(* IEC 61131-3 sources: Lasal-MCP/examples/SampleSource/LASALScreenAdvancedSolution/LASALScreenAdvancedSolution/LASALScreenAdvacnedSolution/Stations/Terminal/HMI/Class/CirleMyIO, 1 file *)

(* ---- CirleMyIO.st ---- *)
(*!
<Class
	Name               = "CirleMyIO"
	Revision           = "0.0"
	RealtimeTask       = "false"
	CyclicTask         = "false"
	BackgroundTask     = "false"
	Sigmatek           = "false"
	OSInterface        = "false"
	HighPriority       = "false"
	Automatic          = "false"
	UpdateMode         = "Prescan"
	SharedCommandTable = "true"
	Objectsize         = "(510,660)">
	<Channels>
		<Server Name="CircleAngle" Visualized="true" Initialize="true" DefValue="3600" WriteProtected="false" Retentive="File"/>
		<Server Name="CircleRadius" Visualized="true" Initialize="true" DefValue="80" WriteProtected="false" Retentive="File"/>
		<Server Name="XPos" Visualized="true" Initialize="true" DefValue="60" WriteProtected="false" Retentive="false"/>
		<Server Name="YPos" Visualized="true" Initialize="true" DefValue="60" WriteProtected="false" Retentive="false"/>
		<Client Name="_Grafix" Required="false" Internal="false"/>
	</Channels>
	<Network Name="CirleMyIO">
		<!-- List of Components in this network -->
		<Components>
			<Object
				Name       = "_base"
				Class      = "_MyIO"
				Position   = "(218,120)"
				Visualized = "true"
				Remotely   = "true">
				<Channels>
					<Server Name="Refresh"/>
					<Server Name="Server0"/>
					<Client Name="Graphic"/>
					<Client Name="Lse"/>
				</Channels>
			</Object>
		</Components>
		<Comments>
		</Comments>
		<!-- List of Connections in this network -->
		<Connections>
			<Connection Source="this.Server0" Destination="_base.Server0" Vertices="(706,210),(534,210),"/>
			<Connection Source="this.Refresh" Destination="_base.Refresh" Vertices="(706,270),(534,270),"/>
			<Connection Source="_base.Lse" Destination="this.Lse" Vertices="(218,210),(38,210),"/>
		</Connections>
		<!-- Headerfiles -->
		<Options>
		</Options>
	</Network>
</Class>
*)
#pragma using _MyIO

CirleMyIO : CLASS
: _MyIO
  //Servers:
	XPos 	: SvrCh_DINT;
	YPos 	: SvrCh_DINT;
	CircleRadius 	: SvrCh_DINT;
	CircleAngle 	: SvrCh_DINT;
  //Clients:
	_Grafix 	: CltChCmd__Grafix;
  //Variables:
		myFocus 	: BOOL;
		TempX 	: _KOORD;
		TempY 	: _KOORD;
  //Functions:
				//! <Function Comment="this method will be called once when the focus will be given to this object" Name="GetFocus"/>
	FUNCTION __CDECL VIRTUAL GLOBAL GetFocus
		VAR_INPUT
			pio 	: ^_IO;			//! <Variable Comment="pointer to _IO information" Name="GetFocus.pio"/>
		END_VAR
		VAR_OUTPUT
			retcode (EAX) 	: _DOIT;			//! <Variable Comment="return _IFAILED if you dont want to get the focus on the other hand _IDLE" Name="GetFocus.retcode"/>
		END_VAR;
				//! <Function Comment="this method is called once when the focus is taken from object" Name="KillFocus"/>
	FUNCTION __CDECL VIRTUAL GLOBAL KillFocus
		VAR_INPUT
			pio 	: ^_IO;			//! <Variable Comment="pointer to _IO information" Name="KillFocus.pio"/>
		END_VAR
		VAR_OUTPUT
			retcode (EAX) 	: _DOIT;			//! <Variable Comment="return always _IDLE because you can&apos;t prevent action" Name="KillFocus.retcode"/>
		END_VAR;
				//! <Function Comment="this method is called everytime when the input is active and a event occured" Name="GetEvent"/>
	FUNCTION __CDECL VIRTUAL GLOBAL GetEvent
		VAR_INPUT
			ped 	: ^_EDITOR;			//! <Variable Comment="pointer to _EDITOR information" Name="GetEvent.ped"/>
			pe 	: ^_EVENT;			//! <Variable Comment="pointer to _EVENT information" Name="GetEvent.pe"/>
		END_VAR
		VAR_OUTPUT
			retcode (EAX) 	: _DOIT;			//! <Variable Comment="for the returnstatement there are 3 different possibilities&#13;&#10;  _IDLE ..... the system should goon like it is (system goes on)&#13;&#10;  _IDIDIT ... i did it (system is ready)&#13;&#10;  _IFAILED .. i tried to do my best, but i failed (system is ready)&#13;&#10;" Name="GetEvent.retcode"/>
		END_VAR;
				//! <Function Comment="this method is called everytime when system wants to redraw the io" Name="Draw"/>
	FUNCTION __CDECL VIRTUAL GLOBAL Draw
		VAR_INPUT
			pio 	: ^_IO;			//! <Variable Comment="pointer to _IO information" Name="Draw.pio"/>
			pr 	: ^_RESULT;			//! <Variable Comment="pointer to _RESULT information" Name="Draw.pr"/>
			pv 	: ^_VARIABLE;			//! <Variable Comment="pointer to io _VARIABLE information" Name="Draw.pv"/>
			input 	: BOOL;			//! <Variable Comment="TRUE it&apos;s an input&#13;&#10;FALSE it&apos;s an output" Name="Draw.input"/>
		END_VAR
		VAR_OUTPUT
			retcode (EAX) 	: _DOIT;			//! <Variable Comment="for the returnstatement there are 3 different possibilities&#13;&#10;  _IDLE ..... the system should goon like it is (system goes on)&#13;&#10;  _IDIDIT ... i did it (system is ready)&#13;&#10;  _IFAILED .. i tried to do my best, but i failed (system is re" Name="Draw.retcode"/>
		END_VAR;
				//! <Function Comment="this method is called everytime when system wants to get data for defined io.&#13;&#10;&#13;&#10;pr ........ &#13;&#10;pio ....... pointer to io information&#13;&#10;pv ........ pointer to io variableinformation&#13;&#10;input ..... TRUE it&apos;s an input / FALSE it&apos;s an output&#13;&#10;&#13;&#10;for the returnstatement there are 3 different possibilities&#13;&#10;_IDLE ..... the system should goon like it is (system goes on)&#13;&#10;_IDIDIT ... i did it (system is ready)&#13;&#10;_IFAILED .. i tried to do my best, but i failed (system is ready)&#13;&#10;&#13;&#10;if you want to do it let&apos;s return _IDIDIT and initialize the  structure _RESULT&#13;&#10;" Name="GetData"/>
	FUNCTION __CDECL VIRTUAL GLOBAL GetData
		VAR_INPUT
			pr 	: ^_RESULT;			//! <Variable Comment="pointer to _RESULT information" Name="GetData.pr"/>
			pio 	: ^_IO;			//! <Variable Comment="pointer to _IO information" Name="GetData.pio"/>
			pv 	: ^_VARIABLE;			//! <Variable Comment="pointer to _VARIABLE information given by LSE" Name="GetData.pv"/>
			input 	: BOOL;			//! <Variable Comment="TRUE it&apos;s an input&#13;&#10;FALSE it&apos;s an output" Name="GetData.input"/>
		END_VAR
		VAR_OUTPUT
			retcode (EAX) 	: _DOIT;			//! <Variable Comment="for the returnstatement there are 3 different possibilities&#13;&#10;  _IDLE ..... the system should goon like it is (system goes on)&#13;&#10;  _IDIDIT ... i did it (system is ready)&#13;&#10;  _IFAILED .. i tried to do my best, but i failed (system is ready)" Name="GetData.retcode"/>
		END_VAR;
  //Tables:
	FUNCTION @STD
		VAR_OUTPUT
			ret_code	: CONFSTATES;
		END_VAR;
	FUNCTION GLOBAL TAB @CT_;
END_CLASS;

#pragma usingLtd _Grafix

FUNCTION __CDECL VIRTUAL GLOBAL CirleMyIO::GetData
	VAR_INPUT
		pr 	: ^_RESULT;
		pio 	: ^_IO;
		pv 	: ^_VARIABLE;
		input 	: BOOL;
	END_VAR
	VAR_OUTPUT
		retcode (EAX) 	: _DOIT;
	END_VAR

  _MyIO::GetData(pr:=pr, pio:=pio, pv:=pv, input:=input);

  pr^.value := to_dint((to_udint(XPos) rol 1) xor (to_udint(YPos)) xor (to_udint(CircleAngle)) xor (to_udint(CircleRadius)));

  retcode := _IDIDIT;

END_FUNCTION

FUNCTION __CDECL VIRTUAL GLOBAL CirleMyIO::Draw
	VAR_INPUT
		pio 	: ^_IO;
		pr 	: ^_RESULT;
		pv 	: ^_VARIABLE;
		input 	: BOOL;
	END_VAR
	VAR_OUTPUT
		retcode (EAX) 	: _DOIT;
	END_VAR
  VAR
  	act   : _NEWSCREEN;
  END_VAR

  _MyIO::Draw(pio:=pio, pr:=pr, pv:=pv, input:=input);

  TempX := pio^.space.xy2.x - (pio^.space.xy2.x - pio^.space.xy1.x) + to_int(XPos) - to_int(CircleRadius / 2);
  TempY := pio^.space.xy2.y - (pio^.space.xy2.y - pio^.space.xy1.y) + to_int(YPos) - to_int(CircleRadius / 2);

  push_screen(#act); // switch over to offscreen
  Graphic.Putimage(#pio^.image, DEFKOORD, DEFKOORD); // display background

  _Grafix.Rectangle(x0:=pio^.space.xy1.x,
                    y0:=pio^.space.xy1.y,
                    x1:=pio^.space.xy2.x,
                    y1:=pio^.space.xy2.y,
                    attrib:= pio^.attrib,
                    color:= pio^.colframe);

   _Grafix.Oval(x0:=TempX + 1,   // Draw circle
                y0:=TempY + 1,
                x1:=TempX + to_int(CircleRadius),
                y1:=TempY + to_int(CircleRadius),
                start:=450,
                bend:=to_int(CircleAngle),
                attrib:=pio^.attrib or T_3D,
                color:=_Grafix.MakeColor(backcolor:=YELLOW, frontcolor:=YELLOW));

  pop_screen(#act); // visible screen switched on
  copy_screen(#act, #pio^.space); // copy image on visible screen

  retcode := _IDIDIT;

END_FUNCTION

FUNCTION __CDECL VIRTUAL GLOBAL CirleMyIO::GetEvent
	VAR_INPUT
		ped 	: ^_EDITOR;
		pe 	: ^_EVENT;
	END_VAR
	VAR_OUTPUT
		retcode (EAX) 	: _DOIT;
	END_VAR

  _MyIO::GetEvent(ped:=ped, pe:=pe);

  retcode := _IDLE;

  if pe^.ftype = _EVENT_HIDMOVE | pe^.ftype = _EVENT_HIDPRESS then

    if ((pe^.dot.x >= ped^.input.io.space.xy1.x + (CircleRadius/2))   &
        (pe^.dot.x <= ped^.input.io.space.xy2.x - (CircleRadius/2)-1) &
        (pe^.dot.y >= ped^.input.io.space.xy1.y + (CircleRadius/2))   &
        (pe^.dot.y <= ped^.input.io.space.xy2.y - (CircleRadius/2)-1))  then

       XPos := pe^.dot.x - ped^.input.io.space.xy1.x;
       YPos := pe^.dot.y - ped^.input.io.space.xy1.y;

       retcode := _IDIDIT;
    end_if;

  end_if;

END_FUNCTION

FUNCTION __CDECL VIRTUAL GLOBAL CirleMyIO::GetFocus
	VAR_INPUT
		pio 	: ^_IO;
	END_VAR
	VAR_OUTPUT
		retcode (EAX) 	: _DOIT;
	END_VAR

  _MyIO::GetFocus(pio:=pio);

  myFocus := TRUE;
  retcode := _IDLE;

END_FUNCTION

FUNCTION __CDECL VIRTUAL GLOBAL CirleMyIO::KillFocus
	VAR_INPUT
    pio 	: ^_IO;
  END_VAR
	VAR_OUTPUT
		retcode (EAX) 	: _DOIT;
	END_VAR

  _MyIO::KillFocus(pio:=pio);

  myFocus := FALSE;
  retcode := _IDLE;

END_FUNCTION
